TEXTLIST TextList_InterConnection
  0 = 'Not Connected'
  1 = 'TriBlender'
  2 = 'Production Line'
  3 = 'Tank'
  4 = 'CIP'
   = ''
END_TEXTLIST

(* stored: Version 1.1.0.1, ProductVersion 3.1.4024.12
   TextList TextList_InterConnection: Id {2e26120c-2bce-47cc-a2fb-42ce357bd332} *)
